DATA_BLOCK "HMI_UPDATE"
TITLE =
VERSION : 0.1


  STRUCT
   HMI_GRAPHIC_TOTAL_1 : DWORD ;	//HMI GRAPHIC TOTAL 1
   HMI_GRAPHIC_TOTAL_2 : DWORD ;	//HMI GRAPHIC TOTAL 1
   HMI_FEED_GRAPHIC : DWORD ;	//HMI GRAPHIC FEED TOTAL 1
   HMI_MOTOR_TOTAL_1 : DWORD ;	//HMI MOTOR TOTAL 1
   HMI_ELEVATOR_PROXS : DWORD ;	//HMI ELEVATOR PROXS
   HMI_FLIPPER_PROXS : DWORD ;	//HMI FLIPPER / TURNTABLE PROXS
   HMI_PUSHER_PROXS : DWORD ;	//HMI PUSHER 9 / PIVOT PROXS
   HMI_FEEDER_PROXS : DWORD ;	//HMI FEEDER PROXS
   HMI_SPARE : DWORD ;	//HMI SPARE
   HMI_FEEDER_GRAPHIC : DWORD ;	//HMI FEEDER GRAPHIC
   HMI_MOTOR_GRAPHIC : DWORD ;	//HMI MOTORGRAPHIC
   HMI_MAIN_PAGE_GRAPHIC : DWORD ;	//HMI MAIN SCREEN GRAPHIC
   HMI_SPARE1 : DWORD ;
   HMI_SPARE2 : DWORD ;
   HMI_SPARE3 : DWORD ;
   HMI_SPARE4 : DWORD ;
   HMI_SPARE5 : DWORD ;
   HMI_SPARE6 : DWORD ;
   HMI_SPARE7 : DWORD ;
   HMI_MOTOR_TOTAL1036 : DWORD ;
   HMI_MOTOR_TOTAL1037 : DWORD ;
   HMI_MOTOR_TOTAL1038 : DWORD ;
   HMI_MOTOR_TOTAL1039 : DWORD ;
   HMI_MOTOR_TOTAL10310 : DWORD ;
  END_STRUCT ;
BEGIN
   HMI_GRAPHIC_TOTAL_1 := DW#16#0;
   HMI_GRAPHIC_TOTAL_2 := DW#16#0;
   HMI_FEED_GRAPHIC := DW#16#0;
   HMI_MOTOR_TOTAL_1 := DW#16#0;
   HMI_ELEVATOR_PROXS := DW#16#0;
   HMI_FLIPPER_PROXS := DW#16#0;
   HMI_PUSHER_PROXS := DW#16#0;
   HMI_FEEDER_PROXS := DW#16#0;
   HMI_SPARE := DW#16#0;
   HMI_FEEDER_GRAPHIC := DW#16#0;
   HMI_MOTOR_GRAPHIC := DW#16#0;
   HMI_MAIN_PAGE_GRAPHIC := DW#16#0;
   HMI_SPARE1 := DW#16#0;
   HMI_SPARE2 := DW#16#0;
   HMI_SPARE3 := DW#16#0;
   HMI_SPARE4 := DW#16#0;
   HMI_SPARE5 := DW#16#0;
   HMI_SPARE6 := DW#16#0;
   HMI_SPARE7 := DW#16#0;
   HMI_MOTOR_TOTAL1036 := DW#16#0;
   HMI_MOTOR_TOTAL1037 := DW#16#0;
   HMI_MOTOR_TOTAL1038 := DW#16#0;
   HMI_MOTOR_TOTAL1039 := DW#16#0;
   HMI_MOTOR_TOTAL10310 := DW#16#0;
END_DATA_BLOCK
